Fanuc KAREL source: KT00908.KL

PROGRAM KT00908
%NOLOCKGROUP
%ENVIRONMENT VECTR
VAR
  P1: POSITION
  P2: POSITION
  OUT: VECTOR
BEGIN
  OUT = ORIENT(P1)
END KT00908
